FUNCTION_BLOCK FB_HMI_Monitoring
VAR_INPUT
END_VAR
VAR_OUTPUT
END_VAR
VAR
END_VAR

END_FUNCTION_BLOCK

(* stored: Version 1.1.0.1, ProductVersion 3.1.4024.15
   POU FB_HMI_Monitoring: Id {77925dff-a4fe-48a9-b80a-5aab27010e3d}, SpecialFunc None *)
